SUBAPPLICATION Uebung_094b2_AX (* Wie Uebung_094b_AX, aber mit explizitem 'nichts ausgewaehlt'-Zustand: AOption_AUI_DEMUX_3 statt _2 - K=1 geht auf DummyGroup (neutraler, wirkungsloser Slot), K=2/3 auf die echten OptionalGroup_001/002. Vermeidet das Problem, welcher Zahlenwert 'Aus' bedeuten soll. *)
  (* Standard: 61499-2; Description: Copyright (c) 2026 Meisterschulen am Ostbahnhof This program and the accompanying materials are made available under the terms of the Eclipse Public License 2.0 which is available at https://www.eclipse.org/legal/epl-2.0/ SPDX-License-Identifier: EPL-2.0 *)
  (* Version 1.0, 2026-10-13, Franz Höpfinger, Meisterschulen am Ostbahnhof, Antwort auf die Rueckfrage, welche Zahlenkonvention (0/1 vs. 1/2) fuer die Dropdown-Werte gelten soll: gar keine Override-Zahlenkonvention noetig, einfach einen eigenen Dummy-Slot im DEMUX reservieren. *)
  PACKAGE Uebungen;
  IMPORT Uebungen::const::UT::DefaultPool::InputNumber_I1;
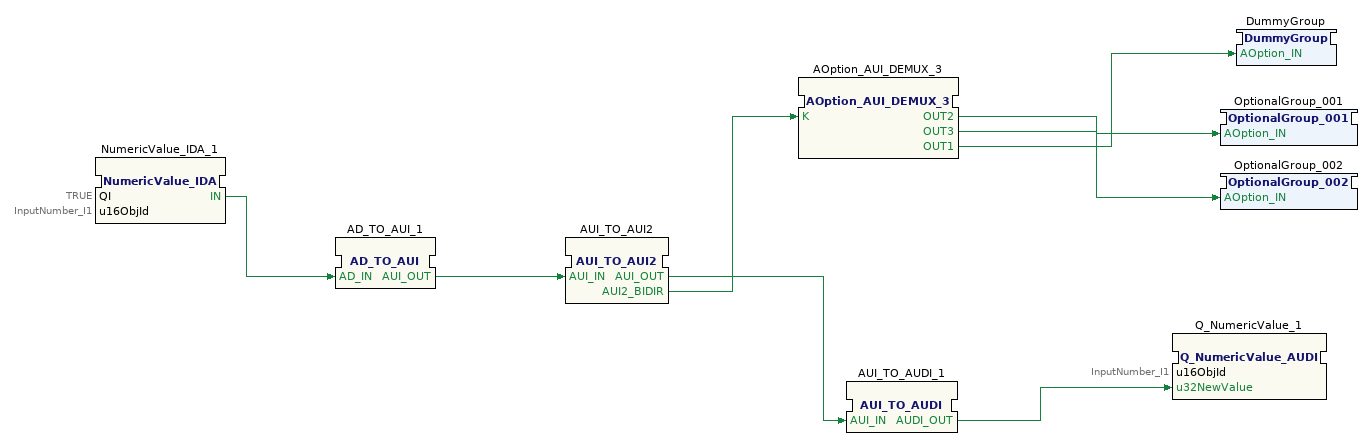
  FBS
    AOption_AUI_DEMUX_3 : Option::selection::AOption_AUI_DEMUX_3;
    NumericValue_IDA_1 : isobus::UT::io::NumericValue::NumericValue_IDA(QI := TRUE, u16ObjId := InputNumber_I1);
    AD_TO_AUI_1 : adapter::conversion::unidirectional::AD_TO_AUI;
    AUI_TO_AUI2 : adapter::conversion::bidirectional::AUI_TO_AUI2;
    AUI_TO_AUDI_1 : adapter::conversion::unidirectional::AUI_TO_AUDI;
    Q_NumericValue_1 : isobus::UT::Q::Q_NumericValue_AUDI(u16ObjId := InputNumber_I1);
  END_FBS
  SUBAPPS
    OptionalGroup_001 : MyLib_AX_Option::sys::OptionalGroup_001;
    OptionalGroup_002 : MyLib_AX_Option::sys::OptionalGroup_002;
    DummyGroup : MyLib_AX_Option::sys::DummyGroup;
  END_SUBAPPS
  ADAPTER_CONNECTIONS
    AOption_AUI_DEMUX_3.OUT2 TO OptionalGroup_001.AOption_IN;
    AOption_AUI_DEMUX_3.OUT3 TO OptionalGroup_002.AOption_IN;
    AOption_AUI_DEMUX_3.OUT1 TO DummyGroup.AOption_IN;
    NumericValue_IDA_1.IN TO AD_TO_AUI_1.AD_IN;
    AUI_TO_AUI2.AUI_OUT TO AUI_TO_AUDI_1.AUI_IN;
    AD_TO_AUI_1.AUI_OUT TO AUI_TO_AUI2.AUI_IN;
    AUI_TO_AUDI_1.AUDI_OUT TO Q_NumericValue_1.u32NewValue;
    AUI_TO_AUI2.AUI2_BIDIR TO AOption_AUI_DEMUX_3.K;
  END_CONNECTIONS
END_SUBAPPLICATION
